{attribute 'no_assign'}
FUNCTION_BLOCK FB_DO_WTURBINE_LD0_WTUR1_TurCtl_st EXTENDS FB_AcsiCommonControllableDataClass
VAR_INPUT
	//stVal: FB_AcsiBATypeEnumerated := (Fc:=ACSI_FC_ST, TrgOp:=ACSI_TrgOp_dchg, bLinkResult:=THIS^.AddDataToContainer(ipData:=stVal));
	stVal: FB_AcsiDATypeTurOp := (Fc:=ACSI_FC_ST, TrgOp:=ACSI_TrgOp_dchg, bLinkResult:=THIS^.AddDataToContainer(ipData:=stVal));
	q: FB_AcsiDATypeQuality := (Fc:=ACSI_FC_ST, TrgOp:=ACSI_TrgOp_qchg, bLinkResult:=THIS^.AddDataToContainer(ipData:=q));
	t: FB_AcsiDATypeTimeStamp := (Fc:=ACSI_FC_ST, bLinkResult:=THIS^.AddDataToContainer(ipData:=t));
	ctlModel: FB_AcsiDATypeCtlModels := (Fc:=ACSI_FC_CF, TrgOp:=ACSI_TrgOp_dchg, eValue:=E_AcsiCtlModels.DirectWithNormalSecurity, bLinkResult:=THIS^.AddDataToContainer(ipData:=ctlModel));
	Cancel: FB_AcsiCDC_Cancel_ENUMERATED := (Fc:=ACSI_FC_CO, bLinkResult:=THIS^.AddDataToContainer(ipData:=Cancel));
	Oper: FB_AcsiCDC_Oper_ENUMERATED := (Fc:=ACSI_FC_CO, bLinkResult:=THIS^.AddDataToContainer(ipData:=Oper));
	SBO: FB_AcsiCDC_SBO := (Fc:=ACSI_FC_CO, bLinkResult:=THIS^.AddDataToContainer(ipData:=SBO));
	
	fbControl: FB_DirectControl := (ipCtrl:=THIS^.AddServerJob(ipEvent:=fbControl, ipCompletion:=fbControl));
END_VAR
VAR
END_VAR

END_FUNCTION_BLOCK

(* stored: Version 1.2.0.0
   POU FB_DO_WTURBINE_LD0_WTUR1_TurCtl_st: Id {8f76b4d8-b90d-4b90-9f49-989661b33e1c}, SpecialFunc None *)
